TYPE ST_BOSCHINDRADRIVECIA402_REF : FB_BOSCHINDRADRIVECIA402_REF;
END_TYPE

(* stored: Version 1.1.0.1, ProductVersion 3.1.4024.15
   DUT ST_BOSCHINDRADRIVECIA402_REF: Id {0a15ad46-8b7e-420d-ad72-82f549a10217} *)
